(* IEC 61131-3 sources: kns-port-domestic/targets/astra/lib/src/POUs/Time/FB_Delay, 3 files *)

(* ---- FB_Delay.decl.st ---- *)
// Назначение: задержка включения и отключения дискретного сигнала — единственный таймер
//             библиотеки (TON, TOF, TP в коде библиотеки не используются). Время берётся из
//             I_TimeSource один раз за вызов; itfTime = 0 — встроенный FB_SystemTime.
//             «Время назад» (ltNow < отметки) перезапускает отсчёт, выход не меняется.
// Автор:      kr0nsch
// Версия:     0.1.0
// Документ:   docs/fb/FB_Delay.md
FUNCTION_BLOCK FB_Delay
VAR_INPUT
    xIn       : BOOL;               // входной сигнал
    tOnDelay  : TIME := T#0S;       // задержка фронта (включения)
    tOffDelay : TIME := T#0S;       // задержка спада (отключения)
    itfTime   : I_TimeSource;       // источник времени; 0 — встроенный fbSysTime
END_VAR
VAR_OUTPUT
    xOut       : BOOL;              // сигнал после задержек
    xTimingOn  : BOOL;              // xIn = TRUE, xOut = FALSE: идёт отсчёт задержки включения
    xTimingOff : BOOL;              // xIn = FALSE, xOut = TRUE: идёт отсчёт задержки отключения
    tRemaining : TIME;              // до смены xOut; T#0S — отсчёта нет
END_VAR
VAR
    fbSysTime : FB_SystemTime;      // запасной источник времени
    ltChange  : LTIME;              // отметка начала отсчёта: смена xIn, первый вызов, Preset, «время назад»
    xInPrev   : BOOL;               // xIn предыдущего вызова
    xRestart  : BOOL := TRUE;       // поставить отметку в ближайшем вызове (первый вызов, Preset)
END_VAR
VAR_TEMP
    ltNow     : LTIME;              // время этого вызова
    ltDelay   : LTIME;              // действующая задержка для текущего xIn
    ltElapsed : LTIME;              // прошло с отметки
END_VAR

(* ---- FB_Delay.impl.st ---- *)
// 1. Время этого вызова — один раз
IF itfTime <> 0 THEN
    ltNow := itfTime.Now();
ELSE
    ltNow := fbSysTime.Now();
END_IF

// 2. Отметка начала отсчёта. Проверка «время назад» — первой: LTIME без знака, и разность
//    ltNow - ltChange при ltNow < ltChange переполнилась бы. Отметка ставится и при смене xIn,
//    в первом вызове и после Preset. После этого шага ltNow >= ltChange.
ltChange := SEL(ltNow < ltChange OR xRestart OR (xIn <> xInPrev), ltChange, ltNow);
xRestart := FALSE;
xInPrev := xIn;

// 3. Задержка для текущего xIn; изменение уставки во время отсчёта действует сразу
// PORT: [types] проверить в Astra.IDE — литералы и преобразования LTIME (C11)
ltDelay := TIME_TO_LTIME(SEL(xIn, tOffDelay, tOnDelay));
ltElapsed := ltNow - ltChange;

// 4. Смена выхода, когда задержка истекла; T#0S — в том же вызове. Если xIn вернулся раньше,
//    xIn = xOut и присваивание ничего не меняет: ожидание отменено
xOut := SEL(ltElapsed >= ltDelay, xOut, xIn);

// 5. Диагностика отсчёта
xTimingOn := xIn AND NOT xOut;
xTimingOff := xOut AND NOT xIn;
IF xIn <> xOut THEN
    // выход не сменился, значит ltElapsed < ltDelay: разность без переполнения
    // PORT: [types] проверить в Astra.IDE — литералы и преобразования LTIME (C11)
    tRemaining := LTIME_TO_TIME(ltDelay - ltElapsed);
ELSE
    tRemaining := T#0S;
END_IF

(* ---- Preset.method.decl.st ---- *)
// Установить выход без задержки (инициализация, выход из подмены, смена режима).
// Отсчёт начнётся заново с ближайшего вызова тела
METHOD PUBLIC Preset
VAR_INPUT
    xValue : BOOL;   // новое значение выхода
END_VAR
